{attribute 'qualified_only'}
{attribute 'strict'}
TYPE E_Prod_Status :
(
	Not_Active := 0,
	Activation_Pending,
	Activation_Pending_Shift, // to shift UTC 
	Active
);
END_TYPE

(* stored: Version 1.1.0.1, ProductVersion 3.1.4024.15
   DUT E_Prod_Status: Id {b75dc2c7-40eb-456a-be1a-10308a6c6645} *)
